INTERFACE ITF_Base

PROPERTY Error : UDINT
GET
END_GET
SET
END_SET
END_PROPERTY

END_INTERFACE

(* stored: Version 1.1.0.1, ProductVersion 3.1.4024.16
   Itf ITF_Base: Id {9d342a4a-d176-4abd-ae0e-b725042d3cc8}
   Property Error: Id {54acd3de-fb7a-427c-a5fb-2211b0a2b32c}
   Get Get: Id {bb431092-a5af-415c-b2c4-e9dc94f83181}
   Set Set: Id {734a7373-d5e4-43d7-9bdb-ab06affef9a4} *)
